Fanuc KAREL source: kb00053.KL

-- PROVISIONAL review KL for V1013-1; original PC SHA256 ae8dcfb4c7326ac04926c8aa899859aff7138af1f8840474211134c2df6f7ac8
-- Incomplete behavior may be omitted. Consult companion uncertainty JSON. Do not deploy.
PROGRAM KB00053
%NOLOCKGROUP
BEGIN
  -- UNRESOLVED_PC offsets 5-15; opcodes 27,31,75
  -- UNRESOLVED_PC offsets 20-24; opcodes 7F
END KB00053
